Staubli VAL3: computeFrame.pgx

program computeFrame(num x_nIndex)
  local num l_nResult
begin

  l_nResult= setFrame(savedata:fFrameItem[x_nIndex].pPointRx[0],savedata:fFrameItem[x_nIndex].pPointRx[1],savedata:fFrameItem[x_nIndex].pPointRx[2],savedata:fFrameItem[x_nIndex].fFrame)
  popUpMsg("坐标系计算完成")
  savedata:libSave()
  delay(0.1)
  if l_nResult<0
    userPageAlert("坐标系示教不成功！请重新示教")
  endIf

end
